INTERFACE I_Maschine

METHOD Start
END_METHOD

METHOD Stop
END_METHOD

METHOD NotausAusloesen
END_METHOD

METHOD NotausZuruecksetzen
END_METHOD

END_INTERFACE

(* stored: Version 1.1.0.1, ProductVersion 3.1.4024.32
   POU I_Maschine: Id {E6B738F9-0A1B-4627-4839-B4C5D6E7F809}, SpecialFunc None
   Method Start: Id {195C0B2D-3E4F-4A5B-6C7D-8E9F0A1B2C3D}
   Method Stop: Id {2A6D1C3E-4F50-4B6C-7D8E-9F0A1B2C3D4E}
   Method NotausAusloesen: Id {3B7E2D4F-5061-4C7D-8E9F-0A1B2C3D4E5F}
   Method NotausZuruecksetzen: Id {4C8F3E50-6172-4D8E-9F0A-1B2C3D4E5F60} *)
